TYPE T_FixtureName : STRING(40); END_TYPE

(* stored: Version 1.1.0.1
   DUT T_FixtureName: Id {2f7c3eb6-52a3-45f2-9733-b5ca1f8fc12d} *)
